{attribute 'qualified_only'}
{attribute 'strict'}
{attribute 'to_string'}
TYPE E_StatusCode :
(
	// The default status.
	STATUS_CODE_UNSET := 0,
	// The Span has been validated by an Application developer or Operator to 
	// have completed successfully.
	STATUS_CODE_OK := 1,
	// The Span contains an error.
	STATUS_CODE_ERROR := 2
) UDINT;
END_TYPE

(* stored: Version 1.1.0.1
   EnumerationTextList E_StatusCode: Id {6c7cce21-2fe4-41e5-8c82-2b54c4e49a98} *)
